(* IEC 61131-3 sources: SRCI_CLIENT_PLC/RobotLibrary/Library/Structures/Telegram/PlcToRob/Cyclic, 1 file *)

(* ---- TelegramPlcToRobCyclicData.st ---- *)
{attribute 'pack_mode' := '1'}
// -------------------------------------------------------------------------
//  SRCI Robot Library
// -------------------------------------------------------------------------
//
//  Object:      TelegramPlcToRobCyclicData
//  Author:      Thorsten Brach
//  Date:        2024-11-30
//
//  Description:
//
//
//  Copyright:
//    (C) 2024 Thorsten Brach. All rights reserved
//             Licensed under the MIT License.
//
//  Disclaimer:
//    This project is provided without any guarantee and can be used for
//    private and commercial purposes. Any use is at the user’s
//    own risk and responsibility.
//
// -------------------------------------------------------------------------
TYPE TelegramPlcToRobCyclicData :
STRUCT
  /// Current Tool
  ToolNo  : BYTE;
  /// Current Frame
  FrameNo : BYTE;
END_STRUCT
END_TYPE
